// TIA Portal V21 export
// export: Created 2026-08-21T20:18:53.9605788Z, ExportSetting None, DisplayName Totally Integrated Automation Portal, DisplayVersion V21, DisplayName STEP 7 Professional, DisplayVersion V21, DisplayName STEP 7 Safety, DisplayVersion V21, DisplayName Tech WebApplication, DisplayVersion V21, DisplayName WinCC Basic/Comfort/Advanced, DisplayVersion V21, DisplayName WinCC Professional, DisplayVersion V21, DisplayName WinCC Unified, DisplayVersion V21
FUNCTION_BLOCK "MTPBinMon_Type1"   // FB16, FBD
{ S7_Optimized_Access := 'TRUE' }
// stored: MemoryReserve 100, SetENOAutomatically false
   VAR_INPUT
      PV { ExternalAccessible := 'False'; ExternalVisible := 'False'; ExternalWritable := 'False'} : Bool;
      PV_QB { ExternalAccessible := 'False'; ExternalVisible := 'False'; ExternalWritable := 'False'} : Bool := true;
      InvPV_In { ExternalAccessible := 'False'; ExternalVisible := 'False'; ExternalWritable := 'False'} : Bool;
   END_VAR
   VAR_OUTPUT
      PV_Out { ExternalAccessible := 'False'; ExternalVisible := 'False'; ExternalWritable := 'False'} : Bool;
      to_Indicate { ExternalAccessible := 'False'; ExternalVisible := 'False'; ExternalWritable := 'False'} : "StruCm";
   END_VAR
   VAR
      DiIn_IDB { ExternalAccessible := 'False'; ExternalVisible := 'False'; ExternalWritable := 'False'} : "DiIn";
      MonDiL_IDB { S7_SetPoint := 'True'} : "MonDiL";
      MTPBinMon_IDB { ExternalVisible := 'False'; S7_SetPoint := 'True'} : "MTPBinMon";
   END_VAR
   VAR_TEMP
      PV_Out_Temp : "DigVal";
      CSF_NOP : "DigVal";
      BadDiIn : "DigVal";
      BadOut : "DigVal";
   END_VAR
   VAR_TEMP   // added for the SCL form of the ladder/FBD networks
      _w1 : Bool;
   END_VAR
BEGIN

REGION Network 1: Analog Input
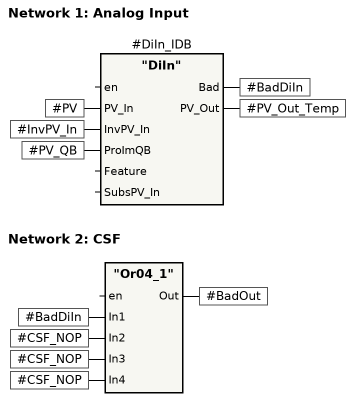
   #DiIn_IDB(PV_In := #PV, InvPV_In := #InvPV_In, ProImQB := #PV_QB, Bad => #BadDiIn, PV_Out => #PV_Out_Temp);   // "DiIn"
END_REGION

REGION Network 2: CSF
   "Or04_1"(In1 := #BadDiIn, In2 := #CSF_NOP, In3 := #CSF_NOP, In4 := #CSF_NOP, Out => #BadOut);
END_REGION

REGION Network 3: MonAnL
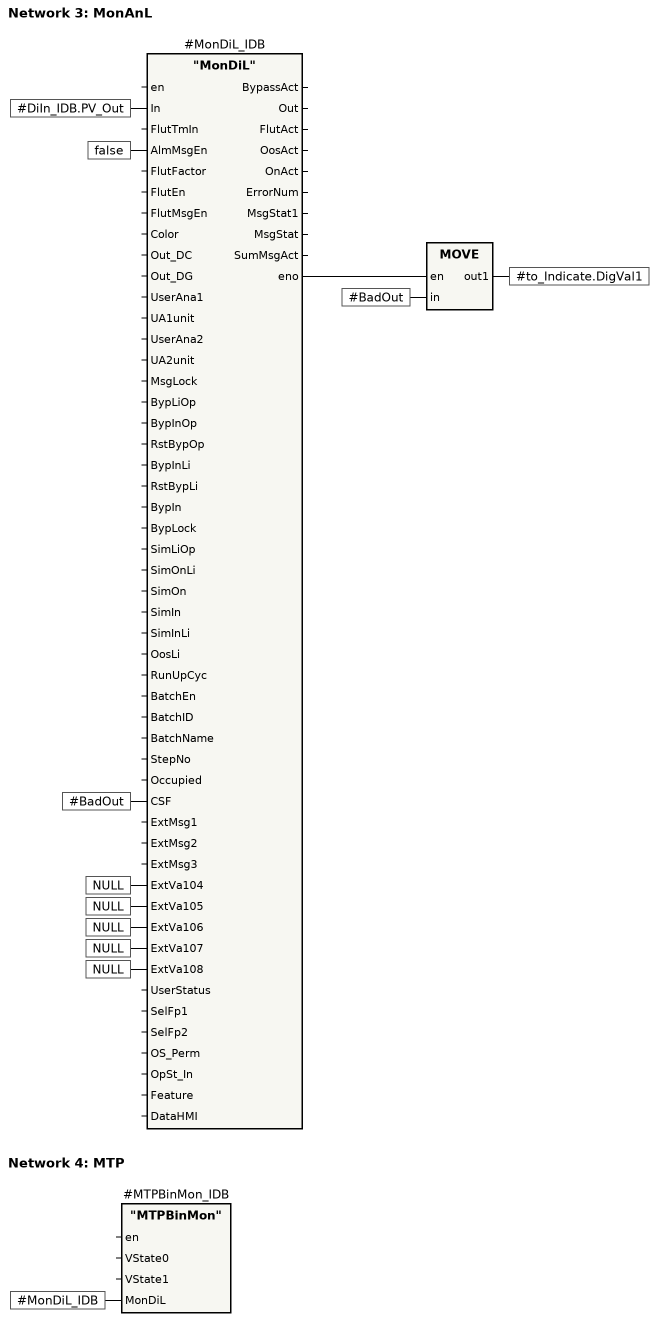
   #MonDiL_IDB(In := #DiIn_IDB.PV_Out,   // "MonDiL"
               AlmMsgEn := false,
               CSF := #BadOut,
               ExtVa104 := NULL,
               ExtVa105 := NULL,
               ExtVa106 := NULL,
               ExtVa107 := NULL,
               ExtVa108 := NULL,
               ENO => #_w1);
   IF #_w1 THEN #to_Indicate.DigVal1 := #BadOut; END_IF;
END_REGION

REGION Network 4: MTP
   #MTPBinMon_IDB(MonDiL := #MonDiL_IDB);   // "MTPBinMon"
END_REGION

REGION Network 5
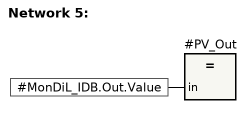
   #PV_Out := #MonDiL_IDB.Out.Value;
END_REGION
END_FUNCTION_BLOCK
